// TIA Portal V20 export
DATA_BLOCK "POS3_0_Messtechnik_DB"   // DB60
// stored: AssignedProDiagFB POS4_0_Prodiag, InstanceOfName POS3_0_Messtechnik, InstanceOfType FB
"POS3_0_Messtechnik"
BEGIN
END_DATA_BLOCK
